(* IEC 61131-3 sources: plc-st-coding-agent/progress/evidence/f14_v14_remaining_20261113/jobs/custom_minimax-m27 (part 4) *)

(* ---- public-medium-02.raw_candidate_03.st ---- *)
TYPE ST_AnalogChannel :
STRUCT
    enable         : BOOL;
    hiLIM          : REAL;
    loLIM          : REAL;
    bipolar        : BOOL;
    measuringMode  : INT;
    retVal         : WORD;
    outputValue    : REAL;
END_STRUCT
END_TYPE;

FUNCTION_BLOCK FB_AnalogBatchProcessing
VAR_INPUT
    count : DINT;
END_VAR
VAR_IN_OUT
    analogValues : ARRAY[*] OF INT;
    channels     : ARRAY[*] OF ST_AnalogChannel;
END_VAR
VAR_OUTPUT
END_VAR
VAR
END_VAR

(*
ENGINEERING_CONTRACT
================================================================================
PUB001: Process 'count' channels starting at each array's lower bound.
        Arrays passed by reference preserve caller-defined bounds.
        Read-only: analogValues elements are never modified.
PUB002: Per-channel conversion based on measuringMode field.
        - Mode 0: Linear scaling using hiLIM/loLIM and bipolar flag.
        - Mode 1: Standard temperature (raw / 10.0).
        - Mode 2: Climatic temperature (raw / 100.0).
        - Invalid mode: retVal=16#8001, outputValue unchanged.
PUB003: Mode 0 linear scaling maps raw 0..27648 (unipolar) or -27648..27648 (bipolar)
        to loLIM..hiLIM range. OutputValue = loLIM + (raw - rawMin) * (hiLIM - loLIM) / range.
PUB004: If hiLIM <= loLIM in mode 0, set retVal=16#8002 and skip conversion.
PUB005: Disabled channels (enable=FALSE) are skipped; retVal and outputValue unchanged.
PUB006: Per-channel retVal WORD status: 16#8001 (invalid mode), 16#8002 (bad range).
PUB007: Same-scan priority: enable→measuringMode→hiLIM/loLIM check→conversion.
PUB008: Temperature output = raw / divisor (10 or 100) as REAL.
--------------------------------------------------------------------------------
*)

VAR
    tmpIndex     : DINT;
    tmpRaw       : INT;
    tmpRawReal   : REAL;
    tmpRange     : REAL;
    tmpOffset    : REAL;
    tmpChannel   : ST_AnalogChannel;
    tmpLower     : DINT;
    tmpUpperAna  : DINT;
    tmpUpperCh   : DINT;
    tmpProcessed : BOOL;
END_VAR

(* CONTRACT_RULES [] *)

tmpLower    := LOWER_BOUND(analogValues, 1);
tmpUpperAna := UPPER_BOUND(analogValues, 1);
tmpUpperCh  := UPPER_BOUND(channels, 1);

FOR tmpIndex := 0 TO (count - 1) DO
    tmpProcessed := FALSE;

    (* Bounds check: skip if index exceeds either array *)
    IF (tmpLower + tmpIndex) <= tmpUpperAna AND (tmpLower + tmpIndex) <= tmpUpperCh THEN
        tmpChannel := channels[tmpLower + tmpIndex];

        (* Skip disabled channels; retain previous outputValue and retVal *)
        IF tmpChannel.enable THEN

    (* Determine conversion based on measuringMode *)
    IF tmpChannel.measuringMode = 0 THEN
        (* Non-temperature linear scaling *)
        IF tmpChannel.hiLIM <= tmpChannel.loLIM THEN
            channels[tmpLower + tmpIndex].retVal := 16#8002;
        ELSE
            tmpRaw       := analogValues[tmpLower + tmpIndex];
            tmpRawReal   := TO_REAL(tmpRaw);
            tmpRange     := tmpChannel.hiLIM - tmpChannel.loLIM;

            IF tmpChannel.bipolar THEN
                (* Map -27648..27648 to loLIM..hiLIM *)
                tmpOffset    := TO_REAL(27648);
                channels[tmpLower + tmpIndex].outputValue := tmpChannel.loLIM +
                    (tmpRawReal + tmpOffset) * tmpRange / TO_REAL(55296);
            ELSE
                (* Map 0..27648 to loLIM..hiLIM *)
                channels[tmpLower + tmpIndex].outputValue := tmpChannel.loLIM +
                    tmpRawReal * tmpRange / TO_REAL(27648);
            END_IF;
            channels[tmpLower + tmpIndex].retVal := 0;
        END_IF;
        tmpProcessed := TRUE;
    ELSIF tmpChannel.measuringMode = 1 THEN
        (* Standard temperature: outputValue = raw / 10 *)
        tmpRaw := analogValues[tmpLower + tmpIndex];
        channels[tmpLower + tmpIndex].outputValue := TO_REAL(tmpRaw) / TO_REAL(10);
        channels[tmpLower + tmpIndex].retVal := 0;
        tmpProcessed := TRUE;
    ELSIF tmpChannel.measuringMode = 2 THEN
        (* Climatic temperature: outputValue = raw / 100 *)
        tmpRaw := analogValues[tmpLower + tmpIndex];
        channels[tmpLower + tmpIndex].outputValue := TO_REAL(tmpRaw) / TO_REAL(100);
        channels[tmpLower + tmpIndex].retVal := 0;
        tmpProcessed := TRUE;
    END_IF;

    (* Invalid measuringMode (not 0, 1, or 2) *)
    IF NOT tmpProcessed THEN
        channels[tmpLower + tmpIndex].retVal := 16#8001;
    END_IF;

    END_IF; (* close outer enable check *)

END_FOR;

END_FUNCTION_BLOCK

(* ---- public-medium-03.candidate_01.st ---- *)
FUNCTION_BLOCK FB_MovingAverage
VAR_INPUT
    cyclicExecution : BOOL;
    trigger         : BOOL;
    value           : LREAL;
    windowSize      : INT;
    reset           : BOOL;
END_VAR
VAR_OUTPUT
    average           : LREAL;
    windowSizeReached : BOOL;
    error             : BOOL;
    status            : WORD;
END_VAR
VAR
    circularBuffer : ARRAY[1..100] OF LREAL;
    bufferIndex    : INT := 1;
    sum             : LREAL := 0.0;
    sampleCount     : INT := 0;
    tmp_triggerPrev : BOOL := FALSE;
END_VAR
VAR_CONSTANT
    STATUS_OK           : WORD := 16#0000;
    STATUS_WINDOW_ERROR : WORD := 16#8200;
END_VAR

(*
ENGINEERING_CONTRACT
===================
Outputs and State Retention:
| Output/State        | Activation                    | Retention                  | Reset/Deactivation       | Same-scan Priority | Units/Boundaries     |
|---------------------|-------------------------------|----------------------------|--------------------------|--------------------| ---------------------|
| average             | New value added (cyclic/trig) | Held until next update     | reset=TRUE clears to 0.0 | cyclic>trigger     | LREAL, windowSize 1-100 |
| windowSizeReached   | sampleCount >= windowSize     | Held TRUE until reset      | reset=TRUE clears FALSE  | N/A                | BOOLEAN             |
| error               | windowSize<1 OR >100          | Held TRUE until valid/reset| reset=TRUE clears FALSE  | N/A                | BOOLEAN             |
| status              | Derived from error state      | Held until state change    | reset=TRUE clears to OK  | N/A                | WORD(16#0000/16#8200) |

Behavior:
- cyclicExecution=TRUE: add value every scan cycle (PUB001)
- trigger rising edge: add one value per press (PUB002)
- cyclicExecution has priority; trigger ignored when cyclic active
- reset clears buffer, sum, count, windowSizeReached (PUB003)
- Invalid windowSize (PUB004) sets error+status and halts processing
- windowSizeReached (PUB005): FALSE until window full, TRUE thereafter
- status codes (PUB006/PUB007): 16#0000=success, 16#8200=window error

First Scan: All VAR initializes to zero/false; no spurious trigger
Boundary: windowSize bounds [1,100] inclusive; strict comparison
)

(* CONTRACT_RULES [] *)

    // Rising edge detection for trigger
    IF trigger AND NOT tmp_triggerPrev THEN
        tmp_triggerPrev := trigger;
        IF NOT reset AND windowSize >= 1 AND windowSize <= 100 THEN
            // Buffer not yet full: add new value
            IF sampleCount < windowSize THEN
                sampleCount := sampleCount + 1;
                circularBuffer[sampleCount] := value;
                sum := sum + value;
                average := sum / TO_LREAL(sampleCount);
                IF sampleCount >= windowSize THEN
                    windowSizeReached := TRUE;
                END_IF;
            ELSE
                // Buffer full: replace oldest value using circular index
                sum := sum - circularBuffer[bufferIndex];
                circularBuffer[bufferIndex] := value;
                sum := sum + value;
                bufferIndex := (bufferIndex MOD windowSize) + 1;
                average := sum / TO_LREAL(windowSize);
            END_IF;
        END_IF;
    ELSE
        tmp_triggerPrev := trigger;
        // Check cyclicExecution on every scan when trigger not rising edge
        IF cyclicExecution AND NOT reset AND windowSize >= 1 AND windowSize <= 100 THEN
            // Buffer not yet full: add new value
            IF sampleCount < windowSize THEN
                sampleCount := sampleCount + 1;
                circularBuffer[sampleCount] := value;
                sum := sum + value;
                average := sum / TO_LREAL(sampleCount);
                IF sampleCount >= windowSize THEN
                    windowSizeReached := TRUE;
                END_IF;
            ELSE
                // Buffer full: replace oldest value using circular index
                sum := sum - circularBuffer[bufferIndex];
                circularBuffer[bufferIndex] := value;
                sum := sum + value;
                bufferIndex := (bufferIndex MOD windowSize) + 1;
                average := sum / TO_LREAL(windowSize);
            END_IF;
        END_IF;
    END_IF;

    // Reset handling - clears all state
    IF reset THEN
        bufferIndex := 1;
        sampleCount := 0;
        sum := 0.0;
        average := 0.0;
        windowSizeReached := FALSE;
        error := FALSE;
        status := STATUS_OK;
    ELSE
        // Validate window size when not resetting
        IF windowSize < 1 OR windowSize > 100 THEN
            error := TRUE;
            status := STATUS_WINDOW_ERROR;
        ELSE
            error := FALSE;
            status := STATUS_OK;
        END_IF;
    END_IF;

END_FUNCTION_BLOCK

(* ---- public-medium-03.candidate_02.st ---- *)
FUNCTION_BLOCK FB_MovingAverage
VAR_INPUT
    cyclicExecution : BOOL;
    trigger         : BOOL;
    value           : LREAL;
    windowSize      : INT;
    reset           : BOOL;
END_VAR
VAR_OUTPUT
    average           : LREAL;
    windowSizeReached : BOOL;
    error             : BOOL;
    status            : WORD;
END_VAR
VAR
    circularBuffer : ARRAY[1..100] OF LREAL;
    bufferIndex    : INT := 1;
    sum             : LREAL := 0.0;
    sampleCount     : INT := 0;
    tmp_triggerPrev : BOOL := FALSE;
END_VAR
VAR
    circularBuffer : ARRAY[1..100] OF LREAL;
    bufferIndex    : INT := 1;
    sum             : LREAL := 0.0;
    sampleCount     : INT := 0;
    tmp_triggerPrev : BOOL := FALSE;
END_VAR

(*
ENGINEERING_CONTRACT
===================
Outputs and State Retention:
| Output/State        | Activation                    | Retention                  | Reset/Deactivation       | Same-scan Priority | Units/Boundaries     |
|---------------------|-------------------------------|----------------------------|--------------------------|--------------------| ---------------------|
| average             | New value added (cyclic/trig) | Held until next update     | reset=TRUE clears to 0.0 | cyclic>trigger     | LREAL, windowSize 1-100 |
| windowSizeReached   | sampleCount >= windowSize     | Held TRUE until reset      | reset=TRUE clears FALSE  | N/A                | BOOLEAN             |
| error               | windowSize<1 OR >100          | Held TRUE until valid/reset| reset=TRUE clears FALSE  | N/A                | BOOLEAN             |
| status              | Derived from error state      | Held until state change    | reset=TRUE clears to OK  | N/A                | WORD(16#0000/16#8200) |

Behavior:
- cyclicExecution=TRUE: add value every scan cycle (PUB001)
- trigger rising edge: add one value per press (PUB002)
- cyclicExecution has priority; trigger ignored when cyclic active
- reset clears buffer, sum, count, windowSizeReached (PUB003)
- Invalid windowSize (PUB004) sets error+status and halts processing
- windowSizeReached (PUB005): FALSE until window full, TRUE thereafter
- status codes (PUB006/PUB007): 16#0000=success, 16#8200=window error

First Scan: All VAR initializes to zero/false; no spurious trigger
Boundary: windowSize bounds [1,100] inclusive; strict comparison
)

(* CONTRACT_RULES [] *)

    // Rising edge detection for trigger
    IF trigger AND NOT tmp_triggerPrev THEN
        tmp_triggerPrev := trigger;
        IF NOT reset AND windowSize >= 1 AND windowSize <= 100 THEN
            // Buffer not yet full: add new value
            IF sampleCount < windowSize THEN
                sampleCount := sampleCount + 1;
                circularBuffer[sampleCount] := value;
                sum := sum + value;
                average := sum / TO_LREAL(sampleCount);
                IF sampleCount >= windowSize THEN
                    windowSizeReached := TRUE;
                END_IF;
            ELSE
                // Buffer full: replace oldest value using circular index
                sum := sum - circularBuffer[bufferIndex];
                circularBuffer[bufferIndex] := value;
                sum := sum + value;
                bufferIndex := (bufferIndex MOD windowSize) + 1;
                average := sum / TO_LREAL(windowSize);
            END_IF;
        END_IF;
    ELSE
        tmp_triggerPrev := trigger;
        // Check cyclicExecution on every scan when trigger not rising edge
        IF cyclicExecution AND NOT reset AND windowSize >= 1 AND windowSize <= 100 THEN
            // Buffer not yet full: add new value
            IF sampleCount < windowSize THEN
                sampleCount := sampleCount + 1;
                circularBuffer[sampleCount] := value;
                sum := sum + value;
                average := sum / TO_LREAL(sampleCount);
                IF sampleCount >= windowSize THEN
                    windowSizeReached := TRUE;
                END_IF;
            ELSE
                // Buffer full: replace oldest value using circular index
                sum := sum - circularBuffer[bufferIndex];
                circularBuffer[bufferIndex] := value;
                sum := sum + value;
                bufferIndex := (bufferIndex MOD windowSize) + 1;
                average := sum / TO_LREAL(windowSize);
            END_IF;
        END_IF;
    END_IF;

    // Reset handling - clears all state
    IF reset THEN
        bufferIndex := 1;
        sampleCount := 0;
        sum := 0.0;
        average := 0.0;
        windowSizeReached := FALSE;
        error := FALSE;
        status := STATUS_OK;
    ELSE
        // Validate window size when not resetting
        IF windowSize < 1 OR windowSize > 100 THEN
            error := TRUE;
            status := STATUS_WINDOW_ERROR;
        ELSE
            error := FALSE;
            status := STATUS_OK;
        END_IF;
    END_IF;

END_FUNCTION_BLOCK

(* ---- public-medium-03.candidate_03.st ---- *)
FUNCTION_BLOCK FB_MovingAverage
VAR_INPUT
    cyclicExecution : BOOL;
    trigger         : BOOL;
    value           : LREAL;
    windowSize      : INT;
    reset           : BOOL;
END_VAR
VAR_OUTPUT
    average           : LREAL;
    windowSizeReached : BOOL;
    error             : BOOL;
    status            : WORD;
END_VAR
VAR
    circularBuffer : ARRAY[1..100] OF LREAL;
    bufferIndex    : INT := 1;
    sum             : LREAL := 0.0;
    sampleCount     : INT := 0;
    tmp_triggerPrev : BOOL := FALSE;
END_VAR

(*
ENGINEERING_CONTRACT
===================
Outputs and State Retention:
| Output/State        | Activation                    | Retention                  | Reset/Deactivation       | Same-scan Priority | Units/Boundaries     |
|---------------------|-------------------------------|----------------------------|--------------------------|--------------------| ---------------------|
| average             | New value added (cyclic/trig) | Held until next update     | reset=TRUE clears to 0.0 | cyclic>trigger     | LREAL, windowSize 1-100 |
| windowSizeReached   | sampleCount >= windowSize     | Held TRUE until reset      | reset=TRUE clears FALSE  | N/A                | BOOLEAN             |
| error               | windowSize<1 OR >100          | Held TRUE until valid/reset| reset=TRUE clears FALSE  | N/A                | BOOLEAN             |
| status              | Derived from error state      | Held until state change    | reset=TRUE clears to OK  | N/A                | WORD(16#0000/16#8200) |

Behavior:
- cyclicExecution=TRUE: add value every scan cycle (PUB001)
- trigger rising edge: add one value per press (PUB002)
- cyclicExecution has priority; trigger ignored when cyclic active
- reset clears buffer, sum, count, windowSizeReached (PUB003)
- Invalid windowSize (PUB004) sets error+status and halts processing
- windowSizeReached (PUB005): FALSE until window full, TRUE thereafter
- status codes (PUB006/PUB007): 16#0000=success, 16#8200=window error

First Scan: All VAR initializes to zero/false; no spurious trigger
Boundary: windowSize bounds [1,100] inclusive; strict comparison
*)

(* CONTRACT_RULES [] *)

    // Rising edge detection for trigger
    IF trigger AND NOT tmp_triggerPrev THEN
        tmp_triggerPrev := trigger;
        IF NOT reset AND windowSize >= 1 AND windowSize <= 100 THEN
            // Buffer not yet full: add new value
            IF sampleCount < windowSize THEN
                sampleCount := sampleCount + 1;
                circularBuffer[sampleCount] := value;
                sum := sum + value;
                average := sum / TO_LREAL(sampleCount);
                IF sampleCount >= windowSize THEN
                    windowSizeReached := TRUE;
                END_IF;
            ELSE
                // Buffer full: replace oldest value using circular index
                sum := sum - circularBuffer[bufferIndex];
                circularBuffer[bufferIndex] := value;
                sum := sum + value;
                bufferIndex := (bufferIndex MOD windowSize) + 1;
                average := sum / TO_LREAL(windowSize);
            END_IF;
        END_IF;
    ELSE
        tmp_triggerPrev := trigger;
        // Check cyclicExecution on every scan when trigger not rising edge
        IF cyclicExecution AND NOT reset AND windowSize >= 1 AND windowSize <= 100 THEN
            // Buffer not yet full: add new value
            IF sampleCount < windowSize THEN
                sampleCount := sampleCount + 1;
                circularBuffer[sampleCount] := value;
                sum := sum + value;
                average := sum / TO_LREAL(sampleCount);
                IF sampleCount >= windowSize THEN
                    windowSizeReached := TRUE;
                END_IF;
            ELSE
                // Buffer full: replace oldest value using circular index
                sum := sum - circularBuffer[bufferIndex];
                circularBuffer[bufferIndex] := value;
                sum := sum + value;
                bufferIndex := (bufferIndex MOD windowSize) + 1;
                average := sum / TO_LREAL(windowSize);
            END_IF;
        END_IF;
    END_IF;

    // Reset handling - clears all state
    IF reset THEN
        bufferIndex := 1;
        sampleCount := 0;
        sum := 0.0;
        average := 0.0;
        windowSizeReached := FALSE;
        error := FALSE;
        status := 16#0000;
    ELSE
        // Validate window size when not resetting
        IF windowSize < 1 OR windowSize > 100 THEN
            error := TRUE;
            status := 16#8200;
        ELSE
            error := FALSE;
            status := 16#0000;
        END_IF;
    END_IF;

END_FUNCTION_BLOCK

(* ---- public-medium-03.candidate_04.st ---- *)
FUNCTION_BLOCK FB_MovingAverage
VAR_INPUT
    cyclicExecution : BOOL;
    trigger         : BOOL;
    value           : LREAL;
    windowSize      : INT;
    reset           : BOOL;
END_VAR
VAR_OUTPUT
    average           : LREAL;
    windowSizeReached : BOOL;
    error             : BOOL;
    status            : WORD;
END_VAR
VAR
    circularBuffer    : ARRAY[1..100] OF LREAL;
    bufferIndex       : INT := 1;
    sum               : LREAL := 0.0;
    sampleCount       : INT := 0;
    tmp_triggerPrev   : BOOL := FALSE;
    tmp_windowSizePrev : INT := 0;
END_VAR

(*
ENGINEERING_CONTRACT
===================
Outputs and State Retention:
| Output/State        | Activation                    | Retention                  | Reset/Deactivation       | Same-scan Priority | Units/Boundaries     |
|---------------------|-------------------------------|----------------------------|--------------------------|--------------------| ---------------------|
| average             | New value added (cyclic/trig) | Held until next update     | reset=TRUE clears to 0.0 | cyclic>trigger     | LREAL, windowSize 1-100 |
| windowSizeReached   | sampleCount >= windowSize     | Held TRUE until reset      | reset=TRUE clears FALSE  | N/A                | BOOLEAN             |
| error               | windowSize<1 OR >100          | Held TRUE until valid/reset| reset=TRUE clears FALSE  | N/A                | BOOLEAN             |
| status              | Derived from error state      | Held until state change    | reset=TRUE clears to OK  | N/A                | WORD(16#0000/16#8200) |

Behavior:
- cyclicExecution=TRUE: add value every scan cycle (PUB001)
- trigger rising edge: add one value per press (PUB002)
- cyclicExecution has priority; trigger ignored when cyclic active
- reset clears buffer, sum, count, windowSizeReached (PUB003)
- Invalid windowSize (PUB004) sets error+status and halts processing
- windowSizeReached (PUB005): FALSE until window full, TRUE thereafter
- status codes (PUB006/PUB007): 16#0000=success, 16#8200=window error

First Scan: All VAR initializes to zero/false; no spurious trigger
Boundary: windowSize bounds [1,100] inclusive; strict comparison
*)

(* CONTRACT_RULES [] *)

    // Detect windowSize change and reset buffer state
    IF windowSize <> tmp_windowSizePrev THEN
        tmp_windowSizePrev := windowSize;
        FOR i := 1 TO 100 DO
            circularBuffer[i] := 0.0;
        END_FOR;
        bufferIndex := 1;
        sampleCount := 0;
        sum := 0.0;
    END_IF;

    // Rising edge detection for trigger takes priority over cyclicExecution
    IF trigger AND NOT tmp_triggerPrev THEN
        tmp_triggerPrev := trigger;
        IF NOT reset AND windowSize >= 1 AND windowSize <= 100 THEN
            // Buffer not yet full: add new value
            IF sampleCount < windowSize THEN
                sampleCount := sampleCount + 1;
                circularBuffer[sampleCount] := value;
                sum := sum + value;
                average := sum / TO_LREAL(sampleCount);
                IF sampleCount >= windowSize THEN
                    windowSizeReached := TRUE;
                END_IF;
            ELSE
                // Buffer full: replace oldest value using circular index
                sum := sum - circularBuffer[bufferIndex];
                circularBuffer[bufferIndex] := value;
                sum := sum + value;
                bufferIndex := (bufferIndex MOD windowSize) + 1;
                average := sum / TO_LREAL(windowSize);
            END_IF;
        END_IF;
    ELSIF cyclicExecution AND NOT tmp_triggerPrev THEN
        tmp_triggerPrev := trigger;
        // cyclicExecution every scan cycle when trigger not active
        IF NOT reset AND windowSize >= 1 AND windowSize <= 100 THEN
            // Buffer not yet full: add new value
            IF sampleCount < windowSize THEN
                sampleCount := sampleCount + 1;
                circularBuffer[sampleCount] := value;
                sum := sum + value;
                average := sum / TO_LREAL(sampleCount);
                IF sampleCount >= windowSize THEN
                    windowSizeReached := TRUE;
                END_IF;
            ELSE
                // Buffer full: replace oldest value using circular index
                sum := sum - circularBuffer[bufferIndex];
                circularBuffer[bufferIndex] := value;
                sum := sum + value;
                bufferIndex := (bufferIndex MOD windowSize) + 1;
                average := sum / TO_LREAL(windowSize);
            END_IF;
        END_IF;
    ELSE
        tmp_triggerPrev := trigger;
    END_IF;

    // Reset handling - clears all state
    IF reset THEN
        bufferIndex := 1;
        sampleCount := 0;
        sum := 0.0;
        average := 0.0;
        windowSizeReached := FALSE;
        error := FALSE;
        status := 16#0000;
    ELSE
        // Validate window size when not resetting
        IF windowSize < 1 OR windowSize > 100 THEN
            error := TRUE;
            status := 16#8200;
        ELSE
            error := FALSE;
            status := 16#0000;
        END_IF;
    END_IF;

END_FUNCTION_BLOCK

(* ---- public-medium-03.patch_base_02.st ---- *)
FUNCTION_BLOCK FB_MovingAverage
VAR_INPUT
    cyclicExecution : BOOL;
    trigger         : BOOL;
    value           : LREAL;
    windowSize      : INT;
    reset           : BOOL;
END_VAR
VAR_OUTPUT
    average           : LREAL;
    windowSizeReached : BOOL;
    error             : BOOL;
    status            : WORD;
END_VAR
VAR
    circularBuffer : ARRAY[1..100] OF LREAL;
    bufferIndex    : INT := 1;
    sum             : LREAL := 0.0;
    sampleCount     : INT := 0;
    tmp_triggerPrev : BOOL := FALSE;
END_VAR
VAR_CONSTANT
    STATUS_OK           : WORD := 16#0000;
    STATUS_WINDOW_ERROR : WORD := 16#8200;
END_VAR

(*
ENGINEERING_CONTRACT
===================
Outputs and State Retention:
| Output/State        | Activation                    | Retention                  | Reset/Deactivation       | Same-scan Priority | Units/Boundaries     |
|---------------------|-------------------------------|----------------------------|--------------------------|--------------------| ---------------------|
| average             | New value added (cyclic/trig) | Held until next update     | reset=TRUE clears to 0.0 | cyclic>trigger     | LREAL, windowSize 1-100 |
| windowSizeReached   | sampleCount >= windowSize     | Held TRUE until reset      | reset=TRUE clears FALSE  | N/A                | BOOLEAN             |
| error               | windowSize<1 OR >100          | Held TRUE until valid/reset| reset=TRUE clears FALSE  | N/A                | BOOLEAN             |
| status              | Derived from error state      | Held until state change    | reset=TRUE clears to OK  | N/A                | WORD(16#0000/16#8200) |

Behavior:
- cyclicExecution=TRUE: add value every scan cycle (PUB001)
- trigger rising edge: add one value per press (PUB002)
- cyclicExecution has priority; trigger ignored when cyclic active
- reset clears buffer, sum, count, windowSizeReached (PUB003)
- Invalid windowSize (PUB004) sets error+status and halts processing
- windowSizeReached (PUB005): FALSE until window full, TRUE thereafter
- status codes (PUB006/PUB007): 16#0000=success, 16#8200=window error

First Scan: All VAR initializes to zero/false; no spurious trigger
Boundary: windowSize bounds [1,100] inclusive; strict comparison
)

(* CONTRACT_RULES [] *)

    // Rising edge detection for trigger
    IF trigger AND NOT tmp_triggerPrev THEN
        tmp_triggerPrev := trigger;
        IF NOT reset AND windowSize >= 1 AND windowSize <= 100 THEN
            // Buffer not yet full: add new value
            IF sampleCount < windowSize THEN
                sampleCount := sampleCount + 1;
                circularBuffer[sampleCount] := value;
                sum := sum + value;
                average := sum / TO_LREAL(sampleCount);
                IF sampleCount >= windowSize THEN
                    windowSizeReached := TRUE;
                END_IF;
            ELSE
                // Buffer full: replace oldest value using circular index
                sum := sum - circularBuffer[bufferIndex];
                circularBuffer[bufferIndex] := value;
                sum := sum + value;
                bufferIndex := (bufferIndex MOD windowSize) + 1;
                average := sum / TO_LREAL(windowSize);
            END_IF;
        END_IF;
    ELSE
        tmp_triggerPrev := trigger;
        // Check cyclicExecution on every scan when trigger not rising edge
        IF cyclicExecution AND NOT reset AND windowSize >= 1 AND windowSize <= 100 THEN
            // Buffer not yet full: add new value
            IF sampleCount < windowSize THEN
                sampleCount := sampleCount + 1;
                circularBuffer[sampleCount] := value;
                sum := sum + value;
                average := sum / TO_LREAL(sampleCount);
                IF sampleCount >= windowSize THEN
                    windowSizeReached := TRUE;
                END_IF;
            ELSE
                // Buffer full: replace oldest value using circular index
                sum := sum - circularBuffer[bufferIndex];
                circularBuffer[bufferIndex] := value;
                sum := sum + value;
                bufferIndex := (bufferIndex MOD windowSize) + 1;
                average := sum / TO_LREAL(windowSize);
            END_IF;
        END_IF;
    END_IF;

    // Reset handling - clears all state
    IF reset THEN
        bufferIndex := 1;
        sampleCount := 0;
        sum := 0.0;
        average := 0.0;
        windowSizeReached := FALSE;
        error := FALSE;
        status := STATUS_OK;
    ELSE
        // Validate window size when not resetting
        IF windowSize < 1 OR windowSize > 100 THEN
            error := TRUE;
            status := STATUS_WINDOW_ERROR;
        ELSE
            error := FALSE;
            status := STATUS_OK;
        END_IF;
    END_IF;

END_FUNCTION_BLOCK

(* ---- public-medium-03.patch_base_03.st ---- *)
FUNCTION_BLOCK FB_MovingAverage
VAR_INPUT
    cyclicExecution : BOOL;
    trigger         : BOOL;
    value           : LREAL;
    windowSize      : INT;
    reset           : BOOL;
END_VAR
VAR_OUTPUT
    average           : LREAL;
    windowSizeReached : BOOL;
    error             : BOOL;
    status            : WORD;
END_VAR
VAR
    circularBuffer : ARRAY[1..100] OF LREAL;
    bufferIndex    : INT := 1;
    sum             : LREAL := 0.0;
    sampleCount     : INT := 0;
    tmp_triggerPrev : BOOL := FALSE;
END_VAR
VAR_CONSTANT
    STATUS_OK           : WORD := 16#0000;
    STATUS_WINDOW_ERROR : WORD := 16#8200;
END_VAR

(*
ENGINEERING_CONTRACT
===================
Outputs and State Retention:
| Output/State        | Activation                    | Retention                  | Reset/Deactivation       | Same-scan Priority | Units/Boundaries     |
|---------------------|-------------------------------|----------------------------|--------------------------|--------------------| ---------------------|
| average             | New value added (cyclic/trig) | Held until next update     | reset=TRUE clears to 0.0 | cyclic>trigger     | LREAL, windowSize 1-100 |
| windowSizeReached   | sampleCount >= windowSize     | Held TRUE until reset      | reset=TRUE clears FALSE  | N/A                | BOOLEAN             |
| error               | windowSize<1 OR >100          | Held TRUE until valid/reset| reset=TRUE clears FALSE  | N/A                | BOOLEAN             |
| status              | Derived from error state      | Held until state change    | reset=TRUE clears to OK  | N/A                | WORD(16#0000/16#8200) |

Behavior:
- cyclicExecution=TRUE: add value every scan cycle (PUB001)
- trigger rising edge: add one value per press (PUB002)
- cyclicExecution has priority; trigger ignored when cyclic active
- reset clears buffer, sum, count, windowSizeReached (PUB003)
- Invalid windowSize (PUB004) sets error+status and halts processing
- windowSizeReached (PUB005): FALSE until window full, TRUE thereafter
- status codes (PUB006/PUB007): 16#0000=success, 16#8200=window error

First Scan: All VAR initializes to zero/false; no spurious trigger
Boundary: windowSize bounds [1,100] inclusive; strict comparison
)

(* CONTRACT_RULES [] *)

    // Rising edge detection for trigger
    IF trigger AND NOT tmp_triggerPrev THEN
        tmp_triggerPrev := trigger;
        IF NOT reset AND windowSize >= 1 AND windowSize <= 100 THEN
            // Buffer not yet full: add new value
            IF sampleCount < windowSize THEN
                sampleCount := sampleCount + 1;
                circularBuffer[sampleCount] := value;
                sum := sum + value;
                average := sum / TO_LREAL(sampleCount);
                IF sampleCount >= windowSize THEN
                    windowSizeReached := TRUE;
                END_IF;
            ELSE
                // Buffer full: replace oldest value using circular index
                sum := sum - circularBuffer[bufferIndex];
                circularBuffer[bufferIndex] := value;
                sum := sum + value;
                bufferIndex := (bufferIndex MOD windowSize) + 1;
                average := sum / TO_LREAL(windowSize);
            END_IF;
        END_IF;
    ELSE
        tmp_triggerPrev := trigger;
        // Check cyclicExecution on every scan when trigger not rising edge
        IF cyclicExecution AND NOT reset AND windowSize >= 1 AND windowSize <= 100 THEN
            // Buffer not yet full: add new value
            IF sampleCount < windowSize THEN
                sampleCount := sampleCount + 1;
                circularBuffer[sampleCount] := value;
                sum := sum + value;
                average := sum / TO_LREAL(sampleCount);
                IF sampleCount >= windowSize THEN
                    windowSizeReached := TRUE;
                END_IF;
            ELSE
                // Buffer full: replace oldest value using circular index
                sum := sum - circularBuffer[bufferIndex];
                circularBuffer[bufferIndex] := value;
                sum := sum + value;
                bufferIndex := (bufferIndex MOD windowSize) + 1;
                average := sum / TO_LREAL(windowSize);
            END_IF;
        END_IF;
    END_IF;

    // Reset handling - clears all state
    IF reset THEN
        bufferIndex := 1;
        sampleCount := 0;
        sum := 0.0;
        average := 0.0;
        windowSizeReached := FALSE;
        error := FALSE;
        status := STATUS_OK;
    ELSE
        // Validate window size when not resetting
        IF windowSize < 1 OR windowSize > 100 THEN
            error := TRUE;
            status := STATUS_WINDOW_ERROR;
        ELSE
            error := FALSE;
            status := STATUS_OK;
        END_IF;
    END_IF;

END_FUNCTION_BLOCK

(* ---- public-medium-03.patch_base_04.st ---- *)
FUNCTION_BLOCK FB_MovingAverage
VAR_INPUT
    cyclicExecution : BOOL;
    trigger         : BOOL;
    value           : LREAL;
    windowSize      : INT;
    reset           : BOOL;
END_VAR
VAR_OUTPUT
    average           : LREAL;
    windowSizeReached : BOOL;
    error             : BOOL;
    status            : WORD;
END_VAR
VAR
    circularBuffer : ARRAY[1..100] OF LREAL;
    bufferIndex    : INT := 1;
    sum             : LREAL := 0.0;
    sampleCount     : INT := 0;
    tmp_triggerPrev : BOOL := FALSE;
END_VAR

(*
ENGINEERING_CONTRACT
===================
Outputs and State Retention:
| Output/State        | Activation                    | Retention                  | Reset/Deactivation       | Same-scan Priority | Units/Boundaries     |
|---------------------|-------------------------------|----------------------------|--------------------------|--------------------| ---------------------|
| average             | New value added (cyclic/trig) | Held until next update     | reset=TRUE clears to 0.0 | cyclic>trigger     | LREAL, windowSize 1-100 |
| windowSizeReached   | sampleCount >= windowSize     | Held TRUE until reset      | reset=TRUE clears FALSE  | N/A                | BOOLEAN             |
| error               | windowSize<1 OR >100          | Held TRUE until valid/reset| reset=TRUE clears FALSE  | N/A                | BOOLEAN             |
| status              | Derived from error state      | Held until state change    | reset=TRUE clears to OK  | N/A                | WORD(16#0000/16#8200) |

Behavior:
- cyclicExecution=TRUE: add value every scan cycle (PUB001)
- trigger rising edge: add one value per press (PUB002)
- cyclicExecution has priority; trigger ignored when cyclic active
- reset clears buffer, sum, count, windowSizeReached (PUB003)
- Invalid windowSize (PUB004) sets error+status and halts processing
- windowSizeReached (PUB005): FALSE until window full, TRUE thereafter
- status codes (PUB006/PUB007): 16#0000=success, 16#8200=window error

First Scan: All VAR initializes to zero/false; no spurious trigger
Boundary: windowSize bounds [1,100] inclusive; strict comparison
*)

(* CONTRACT_RULES [] *)

    // Rising edge detection for trigger
    IF trigger AND NOT tmp_triggerPrev THEN
        tmp_triggerPrev := trigger;
        IF NOT reset AND windowSize >= 1 AND windowSize <= 100 THEN
            // Buffer not yet full: add new value
            IF sampleCount < windowSize THEN
                sampleCount := sampleCount + 1;
                circularBuffer[sampleCount] := value;
                sum := sum + value;
                average := sum / TO_LREAL(sampleCount);
                IF sampleCount >= windowSize THEN
                    windowSizeReached := TRUE;
                END_IF;
            ELSE
                // Buffer full: replace oldest value using circular index
                sum := sum - circularBuffer[bufferIndex];
                circularBuffer[bufferIndex] := value;
                sum := sum + value;
                bufferIndex := (bufferIndex MOD windowSize) + 1;
                average := sum / TO_LREAL(windowSize);
            END_IF;
        END_IF;
    ELSE
        tmp_triggerPrev := trigger;
        // Check cyclicExecution on every scan when trigger not rising edge
        IF cyclicExecution AND NOT reset AND windowSize >= 1 AND windowSize <= 100 THEN
            // Buffer not yet full: add new value
            IF sampleCount < windowSize THEN
                sampleCount := sampleCount + 1;
                circularBuffer[sampleCount] := value;
                sum := sum + value;
                average := sum / TO_LREAL(sampleCount);
                IF sampleCount >= windowSize THEN
                    windowSizeReached := TRUE;
                END_IF;
            ELSE
                // Buffer full: replace oldest value using circular index
                sum := sum - circularBuffer[bufferIndex];
                circularBuffer[bufferIndex] := value;
                sum := sum + value;
                bufferIndex := (bufferIndex MOD windowSize) + 1;
                average := sum / TO_LREAL(windowSize);
            END_IF;
        END_IF;
    END_IF;

    // Reset handling - clears all state
    IF reset THEN
        bufferIndex := 1;
        sampleCount := 0;
        sum := 0.0;
        average := 0.0;
        windowSizeReached := FALSE;
        error := FALSE;
        status := 16#0000;
    ELSE
        // Validate window size when not resetting
        IF windowSize < 1 OR windowSize > 100 THEN
            error := TRUE;
            status := 16#8200;
        ELSE
            error := FALSE;
            status := 16#0000;
        END_IF;
    END_IF;

END_FUNCTION_BLOCK

(* ---- public-medium-03.raw_candidate_01.st ---- *)
FUNCTION_BLOCK FB_MovingAverage
VAR_INPUT
    cyclicExecution : BOOL;
    trigger         : BOOL;
    value           : LREAL;
    windowSize      : INT;
    reset           : BOOL;
END_VAR
VAR_OUTPUT
    average           : LREAL;
    windowSizeReached : BOOL;
    error             : BOOL;
    status            : WORD;
END_VAR
VAR
    circularBuffer : ARRAY[1..100] OF LREAL;
    bufferIndex    : INT := 1;
    sum             : LREAL := 0.0;
    sampleCount     : INT := 0;
    tmp_triggerPrev : BOOL := FALSE;
END_VAR
VAR_CONSTANT
    STATUS_OK           : WORD := 16#0000;
    STATUS_WINDOW_ERROR : WORD := 16#8200;
END_VAR

(*
ENGINEERING_CONTRACT
===================
Outputs and State Retention:
| Output/State        | Activation                    | Retention                  | Reset/Deactivation       | Same-scan Priority | Units/Boundaries     |
|---------------------|-------------------------------|----------------------------|--------------------------|--------------------| ---------------------|
| average             | New value added (cyclic/trig) | Held until next update     | reset=TRUE clears to 0.0 | cyclic>trigger     | LREAL, windowSize 1-100 |
| windowSizeReached   | sampleCount >= windowSize     | Held TRUE until reset      | reset=TRUE clears FALSE  | N/A                | BOOLEAN             |
| error               | windowSize<1 OR >100          | Held TRUE until valid/reset| reset=TRUE clears FALSE  | N/A                | BOOLEAN             |
| status              | Derived from error state      | Held until state change    | reset=TRUE clears to OK  | N/A                | WORD(16#0000/16#8200) |

Behavior:
- cyclicExecution=TRUE: add value every scan cycle (PUB001)
- trigger rising edge: add one value per press (PUB002)
- cyclicExecution has priority; trigger ignored when cyclic active
- reset clears buffer, sum, count, windowSizeReached (PUB003)
- Invalid windowSize (PUB004) sets error+status and halts processing
- windowSizeReached (PUB005): FALSE until window full, TRUE thereafter
- status codes (PUB006/PUB007): 16#0000=success, 16#8200=window error

First Scan: All VAR initializes to zero/false; no spurious trigger
Boundary: windowSize bounds [1,100] inclusive; strict comparison
)

(* CONTRACT_RULES [] *)

    // Rising edge detection for trigger
    IF trigger AND NOT tmp_triggerPrev THEN
        tmp_triggerPrev := trigger;
        IF NOT reset AND windowSize >= 1 AND windowSize <= 100 THEN
            // Buffer not yet full: add new value
            IF sampleCount < windowSize THEN
                sampleCount := sampleCount + 1;
                circularBuffer[sampleCount] := value;
                sum := sum + value;
                average := sum / TO_LREAL(sampleCount);
                IF sampleCount >= windowSize THEN
                    windowSizeReached := TRUE;
                END_IF;
            ELSE
                // Buffer full: replace oldest value using circular index
                sum := sum - circularBuffer[bufferIndex];
                circularBuffer[bufferIndex] := value;
                sum := sum + value;
                bufferIndex := (bufferIndex MOD windowSize) + 1;
                average := sum / TO_LREAL(windowSize);
            END_IF;
        END_IF;
    ELSE
        tmp_triggerPrev := trigger;
        // Check cyclicExecution on every scan when trigger not rising edge
        IF cyclicExecution AND NOT reset AND windowSize >= 1 AND windowSize <= 100 THEN
            // Buffer not yet full: add new value
            IF sampleCount < windowSize THEN
                sampleCount := sampleCount + 1;
                circularBuffer[sampleCount] := value;
                sum := sum + value;
                average := sum / TO_LREAL(sampleCount);
                IF sampleCount >= windowSize THEN
                    windowSizeReached := TRUE;
                END_IF;
            ELSE
                // Buffer full: replace oldest value using circular index
                sum := sum - circularBuffer[bufferIndex];
                circularBuffer[bufferIndex] := value;
                sum := sum + value;
                bufferIndex := (bufferIndex MOD windowSize) + 1;
                average := sum / TO_LREAL(windowSize);
            END_IF;
        END_IF;
    END_IF;

    // Reset handling - clears all state
    IF reset THEN
        bufferIndex := 1;
        sampleCount := 0;
        sum := 0.0;
        average := 0.0;
        windowSizeReached := FALSE;
        error := FALSE;
        status := STATUS_OK;
    ELSE
        // Validate window size when not resetting
        IF windowSize < 1 OR windowSize > 100 THEN
            error := TRUE;
            status := STATUS_WINDOW_ERROR;
        ELSE
            error := FALSE;
            status := STATUS_OK;
        END_IF;
    END_IF;

END_FUNCTION_BLOCK

(* ---- public-medium-03.raw_candidate_02.st ---- *)
FUNCTION_BLOCK FB_MovingAverage
VAR_INPUT
    cyclicExecution : BOOL;
    trigger         : BOOL;
    value           : LREAL;
    windowSize      : INT;
    reset           : BOOL;
END_VAR
VAR_OUTPUT
    average           : LREAL;
    windowSizeReached : BOOL;
    error             : BOOL;
    status            : WORD;
END_VAR
VAR
    circularBuffer : ARRAY[1..100] OF LREAL;
    bufferIndex    : INT := 1;
    sum             : LREAL := 0.0;
    sampleCount     : INT := 0;
    tmp_triggerPrev : BOOL := FALSE;
END_VAR
VAR
    circularBuffer : ARRAY[1..100] OF LREAL;
    bufferIndex    : INT := 1;
    sum             : LREAL := 0.0;
    sampleCount     : INT := 0;
    tmp_triggerPrev : BOOL := FALSE;
END_VAR

(*
ENGINEERING_CONTRACT
===================
Outputs and State Retention:
| Output/State        | Activation                    | Retention                  | Reset/Deactivation       | Same-scan Priority | Units/Boundaries     |
|---------------------|-------------------------------|----------------------------|--------------------------|--------------------| ---------------------|
| average             | New value added (cyclic/trig) | Held until next update     | reset=TRUE clears to 0.0 | cyclic>trigger     | LREAL, windowSize 1-100 |
| windowSizeReached   | sampleCount >= windowSize     | Held TRUE until reset      | reset=TRUE clears FALSE  | N/A                | BOOLEAN             |
| error               | windowSize<1 OR >100          | Held TRUE until valid/reset| reset=TRUE clears FALSE  | N/A                | BOOLEAN             |
| status              | Derived from error state      | Held until state change    | reset=TRUE clears to OK  | N/A                | WORD(16#0000/16#8200) |

Behavior:
- cyclicExecution=TRUE: add value every scan cycle (PUB001)
- trigger rising edge: add one value per press (PUB002)
- cyclicExecution has priority; trigger ignored when cyclic active
- reset clears buffer, sum, count, windowSizeReached (PUB003)
- Invalid windowSize (PUB004) sets error+status and halts processing
- windowSizeReached (PUB005): FALSE until window full, TRUE thereafter
- status codes (PUB006/PUB007): 16#0000=success, 16#8200=window error

First Scan: All VAR initializes to zero/false; no spurious trigger
Boundary: windowSize bounds [1,100] inclusive; strict comparison
)

(* CONTRACT_RULES [] *)

    // Rising edge detection for trigger
    IF trigger AND NOT tmp_triggerPrev THEN
        tmp_triggerPrev := trigger;
        IF NOT reset AND windowSize >= 1 AND windowSize <= 100 THEN
            // Buffer not yet full: add new value
            IF sampleCount < windowSize THEN
                sampleCount := sampleCount + 1;
                circularBuffer[sampleCount] := value;
                sum := sum + value;
                average := sum / TO_LREAL(sampleCount);
                IF sampleCount >= windowSize THEN
                    windowSizeReached := TRUE;
                END_IF;
            ELSE
                // Buffer full: replace oldest value using circular index
                sum := sum - circularBuffer[bufferIndex];
                circularBuffer[bufferIndex] := value;
                sum := sum + value;
                bufferIndex := (bufferIndex MOD windowSize) + 1;
                average := sum / TO_LREAL(windowSize);
            END_IF;
        END_IF;
    ELSE
        tmp_triggerPrev := trigger;
        // Check cyclicExecution on every scan when trigger not rising edge
        IF cyclicExecution AND NOT reset AND windowSize >= 1 AND windowSize <= 100 THEN
            // Buffer not yet full: add new value
            IF sampleCount < windowSize THEN
                sampleCount := sampleCount + 1;
                circularBuffer[sampleCount] := value;
                sum := sum + value;
                average := sum / TO_LREAL(sampleCount);
                IF sampleCount >= windowSize THEN
                    windowSizeReached := TRUE;
                END_IF;
            ELSE
                // Buffer full: replace oldest value using circular index
                sum := sum - circularBuffer[bufferIndex];
                circularBuffer[bufferIndex] := value;
                sum := sum + value;
                bufferIndex := (bufferIndex MOD windowSize) + 1;
                average := sum / TO_LREAL(windowSize);
            END_IF;
        END_IF;
    END_IF;

    // Reset handling - clears all state
    IF reset THEN
        bufferIndex := 1;
        sampleCount := 0;
        sum := 0.0;
        average := 0.0;
        windowSizeReached := FALSE;
        error := FALSE;
        status := STATUS_OK;
    ELSE
        // Validate window size when not resetting
        IF windowSize < 1 OR windowSize > 100 THEN
            error := TRUE;
            status := STATUS_WINDOW_ERROR;
        ELSE
            error := FALSE;
            status := STATUS_OK;
        END_IF;
    END_IF;

END_FUNCTION_BLOCK

(* ---- public-medium-03.raw_candidate_03.st ---- *)
FUNCTION_BLOCK FB_MovingAverage
VAR_INPUT
    cyclicExecution : BOOL;
    trigger         : BOOL;
    value           : LREAL;
    windowSize      : INT;
    reset           : BOOL;
END_VAR
VAR_OUTPUT
    average           : LREAL;
    windowSizeReached : BOOL;
    error             : BOOL;
    status            : WORD;
END_VAR
VAR
    circularBuffer : ARRAY[1..100] OF LREAL;
    bufferIndex    : INT := 1;
    sum             : LREAL := 0.0;
    sampleCount     : INT := 0;
    tmp_triggerPrev : BOOL := FALSE;
END_VAR

(*
ENGINEERING_CONTRACT
===================
Outputs and State Retention:
| Output/State        | Activation                    | Retention                  | Reset/Deactivation       | Same-scan Priority | Units/Boundaries     |
|---------------------|-------------------------------|----------------------------|--------------------------|--------------------| ---------------------|
| average             | New value added (cyclic/trig) | Held until next update     | reset=TRUE clears to 0.0 | cyclic>trigger     | LREAL, windowSize 1-100 |
| windowSizeReached   | sampleCount >= windowSize     | Held TRUE until reset      | reset=TRUE clears FALSE  | N/A                | BOOLEAN             |
| error               | windowSize<1 OR >100          | Held TRUE until valid/reset| reset=TRUE clears FALSE  | N/A                | BOOLEAN             |
| status              | Derived from error state      | Held until state change    | reset=TRUE clears to OK  | N/A                | WORD(16#0000/16#8200) |

Behavior:
- cyclicExecution=TRUE: add value every scan cycle (PUB001)
- trigger rising edge: add one value per press (PUB002)
- cyclicExecution has priority; trigger ignored when cyclic active
- reset clears buffer, sum, count, windowSizeReached (PUB003)
- Invalid windowSize (PUB004) sets error+status and halts processing
- windowSizeReached (PUB005): FALSE until window full, TRUE thereafter
- status codes (PUB006/PUB007): 16#0000=success, 16#8200=window error

First Scan: All VAR initializes to zero/false; no spurious trigger
Boundary: windowSize bounds [1,100] inclusive; strict comparison
*)

(* CONTRACT_RULES [] *)

    // Rising edge detection for trigger
    IF trigger AND NOT tmp_triggerPrev THEN
        tmp_triggerPrev := trigger;
        IF NOT reset AND windowSize >= 1 AND windowSize <= 100 THEN
            // Buffer not yet full: add new value
            IF sampleCount < windowSize THEN
                sampleCount := sampleCount + 1;
                circularBuffer[sampleCount] := value;
                sum := sum + value;
                average := sum / TO_LREAL(sampleCount);
                IF sampleCount >= windowSize THEN
                    windowSizeReached := TRUE;
                END_IF;
            ELSE
                // Buffer full: replace oldest value using circular index
                sum := sum - circularBuffer[bufferIndex];
                circularBuffer[bufferIndex] := value;
                sum := sum + value;
                bufferIndex := (bufferIndex MOD windowSize) + 1;
                average := sum / TO_LREAL(windowSize);
            END_IF;
        END_IF;
    ELSE
        tmp_triggerPrev := trigger;
        // Check cyclicExecution on every scan when trigger not rising edge
        IF cyclicExecution AND NOT reset AND windowSize >= 1 AND windowSize <= 100 THEN
            // Buffer not yet full: add new value
            IF sampleCount < windowSize THEN
                sampleCount := sampleCount + 1;
                circularBuffer[sampleCount] := value;
                sum := sum + value;
                average := sum / TO_LREAL(sampleCount);
                IF sampleCount >= windowSize THEN
                    windowSizeReached := TRUE;
                END_IF;
            ELSE
                // Buffer full: replace oldest value using circular index
                sum := sum - circularBuffer[bufferIndex];
                circularBuffer[bufferIndex] := value;
                sum := sum + value;
                bufferIndex := (bufferIndex MOD windowSize) + 1;
                average := sum / TO_LREAL(windowSize);
            END_IF;
        END_IF;
    END_IF;

    // Reset handling - clears all state
    IF reset THEN
        bufferIndex := 1;
        sampleCount := 0;
        sum := 0.0;
        average := 0.0;
        windowSizeReached := FALSE;
        error := FALSE;
        status := 16#0000;
    ELSE
        // Validate window size when not resetting
        IF windowSize < 1 OR windowSize > 100 THEN
            error := TRUE;
            status := 16#8200;
        ELSE
            error := FALSE;
            status := 16#0000;
        END_IF;
    END_IF;

END_FUNCTION_BLOCK

(* ---- public-medium-03.raw_candidate_04.st ---- *)
FUNCTION_BLOCK FB_MovingAverage
VAR_INPUT
    cyclicExecution : BOOL;
    trigger         : BOOL;
    value           : LREAL;
    windowSize      : INT;
    reset           : BOOL;
END_VAR
VAR_OUTPUT
    average           : LREAL;
    windowSizeReached : BOOL;
    error             : BOOL;
    status            : WORD;
END_VAR
VAR
    circularBuffer    : ARRAY[1..100] OF LREAL;
    bufferIndex       : INT := 1;
    sum               : LREAL := 0.0;
    sampleCount       : INT := 0;
    tmp_triggerPrev   : BOOL := FALSE;
    tmp_windowSizePrev : INT := 0;
END_VAR

(*
ENGINEERING_CONTRACT
===================
Outputs and State Retention:
| Output/State        | Activation                    | Retention                  | Reset/Deactivation       | Same-scan Priority | Units/Boundaries     |
|---------------------|-------------------------------|----------------------------|--------------------------|--------------------| ---------------------|
| average             | New value added (cyclic/trig) | Held until next update     | reset=TRUE clears to 0.0 | cyclic>trigger     | LREAL, windowSize 1-100 |
| windowSizeReached   | sampleCount >= windowSize     | Held TRUE until reset      | reset=TRUE clears FALSE  | N/A                | BOOLEAN             |
| error               | windowSize<1 OR >100          | Held TRUE until valid/reset| reset=TRUE clears FALSE  | N/A                | BOOLEAN             |
| status              | Derived from error state      | Held until state change    | reset=TRUE clears to OK  | N/A                | WORD(16#0000/16#8200) |

Behavior:
- cyclicExecution=TRUE: add value every scan cycle (PUB001)
- trigger rising edge: add one value per press (PUB002)
- cyclicExecution has priority; trigger ignored when cyclic active
- reset clears buffer, sum, count, windowSizeReached (PUB003)
- Invalid windowSize (PUB004) sets error+status and halts processing
- windowSizeReached (PUB005): FALSE until window full, TRUE thereafter
- status codes (PUB006/PUB007): 16#0000=success, 16#8200=window error

First Scan: All VAR initializes to zero/false; no spurious trigger
Boundary: windowSize bounds [1,100] inclusive; strict comparison
*)

(* CONTRACT_RULES [] *)

    // Detect windowSize change and reset buffer state
    IF windowSize <> tmp_windowSizePrev THEN
        tmp_windowSizePrev := windowSize;
        FOR i := 1 TO 100 DO
            circularBuffer[i] := 0.0;
        END_FOR;
        bufferIndex := 1;
        sampleCount := 0;
        sum := 0.0;
    END_IF;

    // Rising edge detection for trigger takes priority over cyclicExecution
    IF trigger AND NOT tmp_triggerPrev THEN
        tmp_triggerPrev := trigger;
        IF NOT reset AND windowSize >= 1 AND windowSize <= 100 THEN
            // Buffer not yet full: add new value
            IF sampleCount < windowSize THEN
                sampleCount := sampleCount + 1;
                circularBuffer[sampleCount] := value;
                sum := sum + value;
                average := sum / TO_LREAL(sampleCount);
                IF sampleCount >= windowSize THEN
                    windowSizeReached := TRUE;
                END_IF;
            ELSE
                // Buffer full: replace oldest value using circular index
                sum := sum - circularBuffer[bufferIndex];
                circularBuffer[bufferIndex] := value;
                sum := sum + value;
                bufferIndex := (bufferIndex MOD windowSize) + 1;
                average := sum / TO_LREAL(windowSize);
            END_IF;
        END_IF;
    ELSIF cyclicExecution AND NOT tmp_triggerPrev THEN
        tmp_triggerPrev := trigger;
        // cyclicExecution every scan cycle when trigger not active
        IF NOT reset AND windowSize >= 1 AND windowSize <= 100 THEN
            // Buffer not yet full: add new value
            IF sampleCount < windowSize THEN
                sampleCount := sampleCount + 1;
                circularBuffer[sampleCount] := value;
                sum := sum + value;
                average := sum / TO_LREAL(sampleCount);
                IF sampleCount >= windowSize THEN
                    windowSizeReached := TRUE;
                END_IF;
            ELSE
                // Buffer full: replace oldest value using circular index
                sum := sum - circularBuffer[bufferIndex];
                circularBuffer[bufferIndex] := value;
                sum := sum + value;
                bufferIndex := (bufferIndex MOD windowSize) + 1;
                average := sum / TO_LREAL(windowSize);
            END_IF;
        END_IF;
    ELSE
        tmp_triggerPrev := trigger;
    END_IF;

    // Reset handling - clears all state
    IF reset THEN
        bufferIndex := 1;
        sampleCount := 0;
        sum := 0.0;
        average := 0.0;
        windowSizeReached := FALSE;
        error := FALSE;
        status := 16#0000;
    ELSE
        // Validate window size when not resetting
        IF windowSize < 1 OR windowSize > 100 THEN
            error := TRUE;
            status := 16#8200;
        ELSE
            error := FALSE;
            status := 16#0000;
        END_IF;
    END_IF;

END_FUNCTION_BLOCK

(* ---- public-medium-04.candidate_01.st ---- *)
FUNCTION_BLOCK FB_TemperatureControl
VAR_INPUT
    TemperatureSensorInput : REAL;
    SetTemperature : REAL;
END_VAR
VAR_OUTPUT
    CurrentTemperature : REAL;
    SetTempDisplay : REAL;
    HeaterStatus : BOOL;
    OverheatProtection : BOOL;
    HeaterOutput : BOOL;
END_VAR
VAR
    OverheatTimer : TON;
    CooldownTimer : TON;
    tmp_SensorFault : BOOL;
END_VAR

(* ENGINEERING_CONTRACT:
 * | Output              | Activation                        | Retention/Hold              | Reset/Deactivation                    | Priority/Scan |
 * |---------------------|------------------------------------|-----------------------------|---------------------------------------|---------------|
 * | CurrentTemperature  | Every scan from sensor             | N/A (combinational read)    | N/A                                   | Same-scan     |
 * | SetTempDisplay      | Every scan from input              | N/A (combinational read)    | N/A                                   | Same-scan     |
 * | HeaterStatus        | Every scan = HeaterOutput          | N/A (combinational mirror)  | N/A                                   | Same-scan     |
 * | HeaterOutput        | Temp < SetTemp AND no fault/protection | Hold while conditions met | Sensor fault OR OverheatProtection OR Temp > SetTemp | Same-scan |
 * | OverheatProtection  | 5s continuous HeaterOutput         | Hold until 3s cooldown done | CooldownTimer.Q (elapsed >= 3s)       | Safety latch  |
 *
 * PUB001: HeaterOutput = (TemperatureSensorInput < SetTemperature) when no faults
 * PUB002, PUB005, PUB006, PUB008: Overheat triggers after TON.Q (elapsed >= 5s) with continuous heater ON
 *         3s cooldown via CooldownTimer before OverheatProtection can clear
 * PUB003: All status outputs updated every scan from current sensor/control state
 * PUB004: Sensor fault (temp < 0 OR temp > 100) disables heater immediately; no hysteresis on fault
 * Units: Temperature [degrees], Time [IEC TON with PT=T#5S/T#3S]
 *)

(* Initialize timers on first scan *)
OverheatTimer(IN := FALSE, PT := T#5S);
CooldownTimer(IN := FALSE, PT := T#3S);

(* PUB004: Sensor fault detection - immediate heater disable *)
tmp_SensorFault := (TemperatureSensorInput < 0.0) OR (TemperatureSensorInput > 100.0);

(* Primary control logic with safety priority *)
IF tmp_SensorFault THEN
    (* PUB004: Sensor fault - disable heater, enter protection state *)
    HeaterOutput := FALSE;
    OverheatProtection := TRUE;
    OverheatTimer(IN := FALSE);
    CooldownTimer(IN := TRUE, PT := T#3S);
    IF CooldownTimer.Q THEN
        OverheatProtection := FALSE;
        CooldownTimer(IN := FALSE);
    END_IF;

ELSIF OverheatProtection THEN
    (* PUB005, PUB008: Overheat protection active - heater forced OFF, cooldown in progress *)
    HeaterOutput := FALSE;
    CooldownTimer(IN := TRUE, PT := T#3S);
    OverheatTimer(IN := FALSE);
    IF CooldownTimer.Q THEN
        OverheatProtection := FALSE;
        CooldownTimer(IN := FALSE);
    END_IF;

ELSE
    (* Normal temperature control *)
    IF TemperatureSensorInput < SetTemperature THEN
        HeaterOutput := TRUE;
    ELSE
        HeaterOutput := FALSE;
    END_IF;

    (* PUB005, PUB006: Overheat protection - track 5s continuous heater operation *)
    IF HeaterOutput THEN
        OverheatTimer(IN := TRUE, PT := T#5S);
        IF OverheatTimer.Q THEN
            (* PUB002, PUB008: Overheat triggered - auto-off heater, start 3s cooldown *)
            OverheatProtection := TRUE;
            HeaterOutput := FALSE;
            OverheatTimer(IN := FALSE);
            CooldownTimer(IN := TRUE, PT := T#3S);
        END_IF;
    ELSE
        OverheatTimer(IN := FALSE);
    END_IF;
END_IF;

(* PUB003: Status display outputs updated every scan *)
CurrentTemperature := TemperatureSensorInput;
SetTempDisplay := SetTemperature;
HeaterStatus := HeaterOutput;
END_FUNCTION_BLOCK

(* CONTRACT_RULES [{"kind": "hold_until_reset", "output": "OverheatProtection", "set_input": null, "reset_input": null}] *)

(* ---- public-medium-04.patch_base_02.st ---- *)
FUNCTION_BLOCK FB_TemperatureControl
VAR_INPUT
    TemperatureSensorInput : REAL;
    SetTemperature : REAL;
END_VAR
VAR_OUTPUT
    CurrentTemperature : REAL;
    SetTempDisplay : REAL;
    HeaterStatus : BOOL;
    OverheatProtection : BOOL;
    HeaterOutput : BOOL;
END_VAR
VAR
    OverheatTimer : TON;
    CooldownTimer : TON;
    tmp_SensorFault : BOOL;
END_VAR

(* ENGINEERING_CONTRACT:
 * | Output              | Activation                        | Retention/Hold              | Reset/Deactivation                    | Priority/Scan |
 * |---------------------|------------------------------------|-----------------------------|---------------------------------------|---------------|
 * | CurrentTemperature  | Every scan from sensor             | N/A (combinational read)    | N/A                                   | Same-scan     |
 * | SetTempDisplay      | Every scan from input              | N/A (combinational read)    | N/A                                   | Same-scan     |
 * | HeaterStatus        | Every scan = HeaterOutput          | N/A (combinational mirror)  | N/A                                   | Same-scan     |
 * | HeaterOutput        | Temp < SetTemp AND no fault/protection | Hold while conditions met | Sensor fault OR OverheatProtection OR Temp > SetTemp | Same-scan |
 * | OverheatProtection  | 5s continuous HeaterOutput         | Hold until 3s cooldown done | CooldownTimer.Q (elapsed >= 3s)       | Safety latch  |
 *
 * PUB001: HeaterOutput = (TemperatureSensorInput < SetTemperature) when no faults
 * PUB002, PUB005, PUB006, PUB008: Overheat triggers after TON.Q (elapsed >= 5s) with continuous heater ON
 *         3s cooldown via CooldownTimer before OverheatProtection can clear
 * PUB003: All status outputs updated every scan from current sensor/control state
 * PUB004: Sensor fault (temp < 0 OR temp > 100) disables heater immediately; no hysteresis on fault
 * Units: Temperature [degrees], Time [IEC TON with PT=T#5S/T#3S]
 *)

(* Initialize timers on first scan *)
OverheatTimer(IN := FALSE, PT := T#5S);
CooldownTimer(IN := FALSE, PT := T#3S);

(* PUB004: Sensor fault detection - immediate heater disable *)
tmp_SensorFault := (TemperatureSensorInput < 0.0) OR (TemperatureSensorInput > 100.0);

(* Primary control logic with safety priority *)
IF tmp_SensorFault THEN
    (* PUB004: Sensor fault - disable heater, enter protection state *)
    HeaterOutput := FALSE;
    OverheatProtection := TRUE;
    OverheatTimer(IN := FALSE);
    CooldownTimer(IN := TRUE, PT := T#3S);
    IF CooldownTimer.Q THEN
        OverheatProtection := FALSE;
        CooldownTimer(IN := FALSE);
    END_IF;

ELSIF OverheatProtection THEN
    (* PUB005, PUB008: Overheat protection active - heater forced OFF, cooldown in progress *)
    HeaterOutput := FALSE;
    CooldownTimer(IN := TRUE, PT := T#3S);
    OverheatTimer(IN := FALSE);
    IF CooldownTimer.Q THEN
        OverheatProtection := FALSE;
        CooldownTimer(IN := FALSE);
    END_IF;

ELSE
    (* Normal temperature control *)
    IF TemperatureSensorInput < SetTemperature THEN
        HeaterOutput := TRUE;
    ELSE
        HeaterOutput := FALSE;
    END_IF;

    (* PUB005, PUB006: Overheat protection - track 5s continuous heater operation *)
    IF HeaterOutput THEN
        OverheatTimer(IN := TRUE, PT := T#5S);
        IF OverheatTimer.Q THEN
            (* PUB002, PUB008: Overheat triggered - auto-off heater, start 3s cooldown *)
            OverheatProtection := TRUE;
            HeaterOutput := FALSE;
            OverheatTimer(IN := FALSE);
            CooldownTimer(IN := TRUE, PT := T#3S);
        END_IF;
    ELSE
        OverheatTimer(IN := FALSE);
    END_IF;
END_IF;

(* PUB003: Status display outputs updated every scan *)
CurrentTemperature := TemperatureSensorInput;
SetTempDisplay := SetTemperature;
HeaterStatus := HeaterOutput;
END_FUNCTION_BLOCK

(* CONTRACT_RULES [{"kind": "hold_until_reset", "output": "OverheatProtection", "set_input": null, "reset_input": null}] *)

(* ---- public-medium-04.patch_base_03.st ---- *)
FUNCTION_BLOCK FB_TemperatureControl
VAR_INPUT
    TemperatureSensorInput : REAL;
    SetTemperature : REAL;
END_VAR
VAR_OUTPUT
    CurrentTemperature : REAL;
    SetTempDisplay : REAL;
    HeaterStatus : BOOL;
    OverheatProtection : BOOL;
    HeaterOutput : BOOL;
END_VAR
VAR
    OverheatTimer : TON;
    CooldownTimer : TON;
    tmp_SensorFault : BOOL;
END_VAR

(* ENGINEERING_CONTRACT:
 * | Output              | Activation                        | Retention/Hold              | Reset/Deactivation                    | Priority/Scan |
 * |---------------------|------------------------------------|-----------------------------|---------------------------------------|---------------|
 * | CurrentTemperature  | Every scan from sensor             | N/A (combinational read)    | N/A                                   | Same-scan     |
 * | SetTempDisplay      | Every scan from input              | N/A (combinational read)    | N/A                                   | Same-scan     |
 * | HeaterStatus        | Every scan = HeaterOutput          | N/A (combinational mirror)  | N/A                                   | Same-scan     |
 * | HeaterOutput        | Temp < SetTemp AND no fault/protection | Hold while conditions met | Sensor fault OR OverheatProtection OR Temp > SetTemp | Same-scan |
 * | OverheatProtection  | 5s continuous HeaterOutput         | Hold until 3s cooldown done | CooldownTimer.Q (elapsed >= 3s)       | Safety latch  |
 *
 * PUB001: HeaterOutput = (TemperatureSensorInput < SetTemperature) when no faults
 * PUB002, PUB005, PUB006, PUB008: Overheat triggers after TON.Q (elapsed >= 5s) with continuous heater ON
 *         3s cooldown via CooldownTimer before OverheatProtection can clear
 * PUB003: All status outputs updated every scan from current sensor/control state
 * PUB004: Sensor fault (temp < 0 OR temp > 100) disables heater immediately; no hysteresis on fault
 * Units: Temperature [degrees], Time [IEC TON with PT=T#5S/T#3S]
 *)

(* Initialize timers on first scan *)
OverheatTimer(IN := FALSE, PT := T#5S);
CooldownTimer(IN := FALSE, PT := T#3S);

(* PUB004: Sensor fault detection - immediate heater disable *)
tmp_SensorFault := (TemperatureSensorInput < 0.0) OR (TemperatureSensorInput > 100.0);

(* Primary control logic with safety priority *)
IF tmp_SensorFault THEN
    (* PUB004: Sensor fault - disable heater, enter protection state *)
    HeaterOutput := FALSE;
    OverheatProtection := TRUE;
    OverheatTimer(IN := FALSE);
    CooldownTimer(IN := TRUE, PT := T#3S);
    IF CooldownTimer.Q THEN
        OverheatProtection := FALSE;
        CooldownTimer(IN := FALSE);
    END_IF;

ELSIF OverheatProtection THEN
    (* PUB005, PUB008: Overheat protection active - heater forced OFF, cooldown in progress *)
    HeaterOutput := FALSE;
    CooldownTimer(IN := TRUE, PT := T#3S);
    OverheatTimer(IN := FALSE);
    IF CooldownTimer.Q THEN
        OverheatProtection := FALSE;
        CooldownTimer(IN := FALSE);
    END_IF;

ELSE
    (* Normal temperature control *)
    IF TemperatureSensorInput < SetTemperature THEN
        HeaterOutput := TRUE;
    ELSE
        HeaterOutput := FALSE;
    END_IF;

    (* PUB005, PUB006: Overheat protection - track 5s continuous heater operation *)
    IF HeaterOutput THEN
        OverheatTimer(IN := TRUE, PT := T#5S);
        IF OverheatTimer.Q THEN
            (* PUB002, PUB008: Overheat triggered - auto-off heater, start 3s cooldown *)
            OverheatProtection := TRUE;
            HeaterOutput := FALSE;
            OverheatTimer(IN := FALSE);
            CooldownTimer(IN := TRUE, PT := T#3S);
        END_IF;
    ELSE
        OverheatTimer(IN := FALSE);
    END_IF;
END_IF;

(* PUB003: Status display outputs updated every scan *)
CurrentTemperature := TemperatureSensorInput;
SetTempDisplay := SetTemperature;
HeaterStatus := HeaterOutput;
END_FUNCTION_BLOCK

(* CONTRACT_RULES [{"kind": "hold_until_reset", "output": "OverheatProtection", "set_input": null, "reset_input": null}] *)

(* ---- public-medium-04.raw_candidate_01.st ---- *)
FUNCTION_BLOCK FB_TemperatureControl
VAR_INPUT
    TemperatureSensorInput : REAL;
    SetTemperature : REAL;
END_VAR
VAR_OUTPUT
    CurrentTemperature : REAL;
    SetTempDisplay : REAL;
    HeaterStatus : BOOL;
    OverheatProtection : BOOL;
    HeaterOutput : BOOL;
END_VAR
VAR
    OverheatTimer : TON;
    CooldownTimer : TON;
    tmp_SensorFault : BOOL;
END_VAR

(* ENGINEERING_CONTRACT:
 * | Output              | Activation                        | Retention/Hold              | Reset/Deactivation                    | Priority/Scan |
 * |---------------------|------------------------------------|-----------------------------|---------------------------------------|---------------|
 * | CurrentTemperature  | Every scan from sensor             | N/A (combinational read)    | N/A                                   | Same-scan     |
 * | SetTempDisplay      | Every scan from input              | N/A (combinational read)    | N/A                                   | Same-scan     |
 * | HeaterStatus        | Every scan = HeaterOutput          | N/A (combinational mirror)  | N/A                                   | Same-scan     |
 * | HeaterOutput        | Temp < SetTemp AND no fault/protection | Hold while conditions met | Sensor fault OR OverheatProtection OR Temp > SetTemp | Same-scan |
 * | OverheatProtection  | 5s continuous HeaterOutput         | Hold until 3s cooldown done | CooldownTimer.Q (elapsed >= 3s)       | Safety latch  |
 *
 * PUB001: HeaterOutput = (TemperatureSensorInput < SetTemperature) when no faults
 * PUB002, PUB005, PUB006, PUB008: Overheat triggers after TON.Q (elapsed >= 5s) with continuous heater ON
 *         3s cooldown via CooldownTimer before OverheatProtection can clear
 * PUB003: All status outputs updated every scan from current sensor/control state
 * PUB004: Sensor fault (temp < 0 OR temp > 100) disables heater immediately; no hysteresis on fault
 * Units: Temperature [degrees], Time [IEC TON with PT=T#5S/T#3S]
 *)

(* Initialize timers on first scan *)
OverheatTimer(IN := FALSE, PT := T#5S);
CooldownTimer(IN := FALSE, PT := T#3S);

(* PUB004: Sensor fault detection - immediate heater disable *)
tmp_SensorFault := (TemperatureSensorInput < 0.0) OR (TemperatureSensorInput > 100.0);

(* Primary control logic with safety priority *)
IF tmp_SensorFault THEN
    (* PUB004: Sensor fault - disable heater, enter protection state *)
    HeaterOutput := FALSE;
    OverheatProtection := TRUE;
    OverheatTimer(IN := FALSE);
    CooldownTimer(IN := TRUE, PT := T#3S);
    IF CooldownTimer.Q THEN
        OverheatProtection := FALSE;
        CooldownTimer(IN := FALSE);
    END_IF;

ELSIF OverheatProtection THEN
    (* PUB005, PUB008: Overheat protection active - heater forced OFF, cooldown in progress *)
    HeaterOutput := FALSE;
    CooldownTimer(IN := TRUE, PT := T#3S);
    OverheatTimer(IN := FALSE);
    IF CooldownTimer.Q THEN
        OverheatProtection := FALSE;
        CooldownTimer(IN := FALSE);
    END_IF;

ELSE
    (* Normal temperature control *)
    IF TemperatureSensorInput < SetTemperature THEN
        HeaterOutput := TRUE;
    ELSE
        HeaterOutput := FALSE;
    END_IF;

    (* PUB005, PUB006: Overheat protection - track 5s continuous heater operation *)
    IF HeaterOutput THEN
        OverheatTimer(IN := TRUE, PT := T#5S);
        IF OverheatTimer.Q THEN
            (* PUB002, PUB008: Overheat triggered - auto-off heater, start 3s cooldown *)
            OverheatProtection := TRUE;
            HeaterOutput := FALSE;
            OverheatTimer(IN := FALSE);
            CooldownTimer(IN := TRUE, PT := T#3S);
        END_IF;
    ELSE
        OverheatTimer(IN := FALSE);
    END_IF;
END_IF;

(* PUB003: Status display outputs updated every scan *)
CurrentTemperature := TemperatureSensorInput;
SetTempDisplay := SetTemperature;
HeaterStatus := HeaterOutput;
END_FUNCTION_BLOCK

(* CONTRACT_RULES [{"kind": "hold_until_reset", "output": "OverheatProtection", "set_input": null, "reset_input": null}] *)

(* ---- public-medium-05.candidate_01.st ---- *)
(* ENGINEERING_CONTRACT
 * =============================================================================
 * Mode Switching (PUB001): Mode=0 manual, Mode=1 automatic. Output state on
 *   mode transition: both Motor outputs cleared, CompletionLight cleared.
 *   Transition detected via rising edge on Mode input variable.
 * Manual Mode (PUB002/PUB003):
 *   - Activation: Mode=0
 *   - Retention: MotorForward holds while ForwardButton=1 AND ReverseButton=0
 *   - Retention: MotorReverse holds while ReverseButton=1 AND ForwardButton=0
 *   - Deactivation: both cleared on any of: ForwardButton=0, ReverseButton=0,
 *     forward+reverse both asserted (interlock drops both), or Mode→1
 *   - Units: combinational, no timer
 * Automatic Mode (PUB004-PUB008):
 *   - Scan behavior: edge-sensitive state machine evaluated every scan
 *   - STATION_A activation: SensorA=TRUE AND State=IDLE
 *   - STATION_B activation: SensorB=TRUE AND State=MOVING_TO_B
 *   - STATION_C activation: SensorC=TRUE AND State=MOVING_TO_C
 *   - MotorForward activation: (State=IDLE AND SensorA=TRUE→ButtonA=TRUE)
 *     OR (State=STATION_A AND ButtonA=TRUE) OR (State=STATION_B AND ButtonB=TRUE)
 *   - MotorForward deactivation: on SensorB (→STATION_B) or SensorC (→STATION_C)
 *   - CompletionLight activation: SensorC=TRUE AND ButtonC=TRUE AND State=STATION_C
 *   - CompletionLight retention: holds until SensorC=FALSE (product removed)
 *   - CompletionLight deactivation: SensorC=FALSE transitions to IDLE
 *   - IDLE reset: State=IDLE when no product detected at any station
 *   - Units: boolean states, no timers
 * Same-scan priority: manual overrides automatic (Mode check first). Within
 *   automatic, state transition clears prior MotorForward before next sensor
 *   evaluation; CompletionLight set after Mode/state checks finalized.
 * Physical interlock: Pub002 prohibits MotorForward AND MotorReverse together.
 * =============================================================================
 *)

(* CONTRACT_RULES [] *)

FUNCTION_BLOCK ProductionLineControl
VAR_INPUT
    Mode            : BOOL;  (* 0=manual, 1=automatic *)
    ForwardButton   : BOOL;
    ReverseButton   : BOOL;
    SensorA         : BOOL;
    SensorB         : BOOL;
    SensorC         : BOOL;
    ButtonA         : BOOL;
    ButtonB         : BOOL;
    ButtonC         : BOOL;
END_VAR
VAR_OUTPUT
    MotorForward    : BOOL;
    MotorReverse    : BOOL;
    CompletionLight : BOOL;
END_VAR
VAR
    State           : INT;  (* 0=IDLE, 1=STATION_A, 2=MOVING_TO_B, 3=STATION_B,
                                4=MOVING_TO_C, 5=STATION_C *)
    tmp_PreviousMode : BOOL;
    tmp_ModeRising   : BOOL;
END_VAR

    (* Constants for state identification *)
    CONST
        IDLE         : INT := 0;
        STATION_A    : INT := 1;
        MOVING_TO_B  : INT := 2;
        STATION_B    : INT := 3;
        MOVING_TO_C  : INT := 4;
        STATION_C    : INT := 5;
    END_CONST

    (* Detect mode transition for reset behavior *)
    tmp_ModeRising := Mode AND NOT tmp_PreviousMode;
    tmp_PreviousMode := Mode;

    (* Reset outputs on mode entry into automatic *)
    IF tmp_ModeRising THEN
        MotorForward    := FALSE;
        MotorReverse    := FALSE;
        CompletionLight := FALSE;
    END_IF;

    (* Mode-based operation dispatch *)
    IF Mode = FALSE THEN
        (* Manual Mode (PUB002/PUB003) *)
        (* Interlock: forward and reverse cannot be energized together *)
        IF ForwardButton AND NOT ReverseButton THEN
            MotorForward := TRUE;
            MotorReverse := FALSE;
        ELSIF ReverseButton AND NOT ForwardButton THEN
            MotorForward := FALSE;
            MotorReverse := TRUE;
        ELSE
            MotorForward := FALSE;
            MotorReverse := FALSE;
        END_IF;
    ELSE
        (* Automatic Mode (PUB004-PUB008) *)
        MotorForward    := FALSE;
        MotorReverse    := FALSE;

        (* State machine evaluation *)
        CASE State OF
            IDLE :
                (* Wait for product at Workstation A *)
                IF SensorA THEN
                    State := STATION_A;
                END_IF;

            STATION_A :
                (* Product at Workstation A, wait for ButtonA *)
                IF ButtonA THEN
                    MotorForward := TRUE;
                    State := MOVING_TO_B;
                END_IF;
                (* Fallback: if product leaves A unexpectedly, return to IDLE *)
                IF NOT SensorA THEN
                    State := IDLE;
                END_IF;

            MOVING_TO_B :
                (* Motor running forward, wait for SensorB *)
                MotorForward := TRUE;
                IF SensorB THEN
                    MotorForward := FALSE;
                    State := STATION_B;
                END_IF;

            STATION_B :
                (* Product at Workstation B, wait for ButtonB *)
                IF ButtonB THEN
                    MotorForward := TRUE;
                    State := MOVING_TO_C;
                END_IF;
                (* Fallback: if product leaves B unexpectedly, return to IDLE *)
                IF NOT SensorB THEN
                    State := IDLE;
                END_IF;

            MOVING_TO_C :
                (* Motor running forward, wait for SensorC *)
                MotorForward := TRUE;
                IF SensorC THEN
                    MotorForward := FALSE;
                    State := STATION_C;
                END_IF;

            STATION_C :
                (* Product at Workstation C, wait for ButtonC, then product removal *)
                IF ButtonC THEN
                    CompletionLight := TRUE;
                END_IF;
                (* Product taken away: light off, return to IDLE *)
                IF NOT SensorC THEN
                    CompletionLight := FALSE;
                    State := IDLE;
                END_IF;

        END_CASE;
    END_IF;

END_FUNCTION_BLOCK

(* ---- public-medium-05.candidate_02.st ---- *)
TYPE ProductionState : INT (
    IDLE := 0,
    STATION_A := 1,
    MOVING_TO_B := 2,
    STATION_B := 3,
    MOVING_TO_C := 4,
    STATION_C := 5
);
END_TYPE;

(* ENGINEERING_CONTRACT
 * =============================================================================
 * Mode Switching (PUB001): Mode=0 manual, Mode=1 automatic. Output state on
 *   mode transition: both Motor outputs cleared, CompletionLight cleared.
 *   Transition detected via rising edge on Mode input variable.
 * Manual Mode (PUB002/PUB003):
 *   - Activation: Mode=0
 *   - Retention: MotorForward holds while ForwardButton=1 AND ReverseButton=0
 *   - Retention: MotorReverse holds while ReverseButton=1 AND ForwardButton=0
 *   - Deactivation: both cleared on any of: ForwardButton=0, ReverseButton=0,
 *     forward+reverse both asserted (interlock drops both), or Mode→1
 *   - Units: combinational, no timer
 * Automatic Mode (PUB004-PUB008):
 *   - Scan behavior: edge-sensitive state machine evaluated every scan
 *   - STATION_A activation: SensorA=TRUE AND State=IDLE
 *   - STATION_B activation: SensorB=TRUE AND State=MOVING_TO_B
 *   - STATION_C activation: SensorC=TRUE AND State=MOVING_TO_C
 *   - MotorForward activation: (State=IDLE AND SensorA=TRUE→ButtonA=TRUE)
 *     OR (State=STATION_A AND ButtonA=TRUE) OR (State=STATION_B AND ButtonB=TRUE)
 *   - MotorForward deactivation: on SensorB (→STATION_B) or SensorC (→STATION_C)
 *   - CompletionLight activation: SensorC=TRUE AND ButtonC=TRUE AND State=STATION_C
 *   - CompletionLight retention: holds until SensorC=FALSE (product removed)
 *   - CompletionLight deactivation: SensorC=FALSE transitions to IDLE
 *   - IDLE reset: State=IDLE when no product detected at any station
 *   - Units: boolean states, no timers
 * Same-scan priority: manual overrides automatic (Mode check first). Within
 *   automatic, state transition clears prior MotorForward before next sensor
 *   evaluation; CompletionLight set after Mode/state checks finalized.
 * Physical interlock: Pub002 prohibits MotorForward AND MotorReverse together.
 * =============================================================================
 *)

(* CONTRACT_RULES [] *)

FUNCTION_BLOCK ProductionLineControl
VAR_INPUT
    Mode            : BOOL;  (* 0=manual, 1=automatic *)
    ForwardButton   : BOOL;
    ReverseButton   : BOOL;
    SensorA         : BOOL;
    SensorB         : BOOL;
    SensorC         : BOOL;
    ButtonA         : BOOL;
    ButtonB         : BOOL;
    ButtonC         : BOOL;
END_VAR
VAR_OUTPUT
    MotorForward    : BOOL;
    MotorReverse    : BOOL;
    CompletionLight : BOOL;
END_VAR
VAR
    State           : INT;  (* 0=IDLE, 1=STATION_A, 2=MOVING_TO_B, 3=STATION_B,
                                4=MOVING_TO_C, 5=STATION_C *)
    tmp_PreviousMode : BOOL;
    tmp_ModeRising   : BOOL;
END_VAR

    (* Constants for state identification *)
    (* Detect mode transition for reset behavior *)
    tmp_ModeRising := Mode AND NOT tmp_PreviousMode;
    tmp_PreviousMode := Mode;

    (* Reset outputs on mode entry into automatic *)
    IF tmp_ModeRising THEN
        MotorForward    := FALSE;
        MotorReverse    := FALSE;
        CompletionLight := FALSE;
    END_IF;

    (* Mode-based operation dispatch *)
    IF Mode = FALSE THEN
        (* Manual Mode (PUB002/PUB003) *)
        (* Interlock: forward and reverse cannot be energized together *)
        IF ForwardButton AND NOT ReverseButton THEN
            MotorForward := TRUE;
            MotorReverse := FALSE;
        ELSIF ReverseButton AND NOT ForwardButton THEN
            MotorForward := FALSE;
            MotorReverse := TRUE;
        ELSE
            MotorForward := FALSE;
            MotorReverse := FALSE;
        END_IF;
    ELSE
        (* Automatic Mode (PUB004-PUB008) *)
        MotorForward    := FALSE;
        MotorReverse    := FALSE;

        (* State machine evaluation *)
        CASE State OF
            IDLE :
                (* Wait for product at Workstation A *)
                IF SensorA THEN
                    State := STATION_A;
                END_IF;

            STATION_A :
                (* Product at Workstation A, wait for ButtonA *)
                IF ButtonA THEN
                    MotorForward := TRUE;
                    State := MOVING_TO_B;
                END_IF;
                (* Fallback: if product leaves A unexpectedly, return to IDLE *)
                IF NOT SensorA THEN
                    State := IDLE;
                END_IF;

            MOVING_TO_B :
                (* Motor running forward, wait for SensorB *)
                MotorForward := TRUE;
                IF SensorB THEN
                    MotorForward := FALSE;
                    State := STATION_B;
                END_IF;

            STATION_B :
                (* Product at Workstation B, wait for ButtonB *)
                IF ButtonB THEN
                    MotorForward := TRUE;
                    State := MOVING_TO_C;
                END_IF;
                (* Fallback: if product leaves B unexpectedly, return to IDLE *)
                IF NOT SensorB THEN
                    State := IDLE;
                END_IF;

            MOVING_TO_C :
                (* Motor running forward, wait for SensorC *)
                MotorForward := TRUE;
                IF SensorC THEN
                    MotorForward := FALSE;
                    State := STATION_C;
                END_IF;

            STATION_C :
                (* Product at Workstation C, wait for ButtonC, then product removal *)
                IF ButtonC THEN
                    CompletionLight := TRUE;
                END_IF;
                (* Product taken away: light off, return to IDLE *)
                IF NOT SensorC THEN
                    CompletionLight := FALSE;
                    State := IDLE;
                END_IF;

        END_CASE;
    END_IF;

END_FUNCTION_BLOCK

(* ---- public-medium-05.candidate_03.st ---- *)
CONST
    IDLE         : INT := 0;
    STATION_A    : INT := 1;
    MOVING_TO_B  : INT := 2;
    STATION_B    : INT := 3;
    MOVING_TO_C  : INT := 4;
    STATION_C    : INT := 5;
END_CONST

(* ENGINEERING_CONTRACT
 * =============================================================================
 * Mode Switching (PUB001): Mode=0 manual, Mode=1 automatic. Output state on
 *   mode transition: both Motor outputs cleared, CompletionLight cleared.
 *   Transition detected via rising edge on Mode input variable.
 * Manual Mode (PUB002/PUB003):
 *   - Activation: Mode=0
 *   - Retention: MotorForward holds while ForwardButton=1 AND ReverseButton=0
 *   - Retention: MotorReverse holds while ReverseButton=1 AND ForwardButton=0
 *   - Deactivation: both cleared on any of: ForwardButton=0, ReverseButton=0,
 *     forward+reverse both asserted (interlock drops both), or Mode→1
 *   - Units: combinational, no timer
 * Automatic Mode (PUB004-PUB008):
 *   - Scan behavior: edge-sensitive state machine evaluated every scan
 *   - STATION_A activation: SensorA=TRUE AND State=IDLE
 *   - STATION_B activation: SensorB=TRUE AND State=MOVING_TO_B
 *   - STATION_C activation: SensorC=TRUE AND State=MOVING_TO_C
 *   - MotorForward activation: (State=IDLE AND SensorA=TRUE→ButtonA=TRUE)
 *     OR (State=STATION_A AND ButtonA=TRUE) OR (State=STATION_B AND ButtonB=TRUE)
 *   - MotorForward deactivation: on SensorB (→STATION_B) or SensorC (→STATION_C)
 *   - CompletionLight activation: SensorC=TRUE AND ButtonC=TRUE AND State=STATION_C
 *   - CompletionLight retention: holds until SensorC=FALSE (product removed)
 *   - CompletionLight deactivation: SensorC=FALSE transitions to IDLE
 *   - IDLE reset: State=IDLE when no product detected at any station
 *   - Units: boolean states, no timers
 * Same-scan priority: manual overrides automatic (Mode check first). Within
 *   automatic, state transition clears prior MotorForward before next sensor
 *   evaluation; CompletionLight set after Mode/state checks finalized.
 * Physical interlock: Pub002 prohibits MotorForward AND MotorReverse together.
 * =============================================================================
 *)

(* CONTRACT_RULES [] *)

FUNCTION_BLOCK ProductionLineControl
VAR_INPUT
    Mode            : BOOL;  (* 0=manual, 1=automatic *)
    ForwardButton   : BOOL;
    ReverseButton   : BOOL;
    SensorA         : BOOL;
    SensorB         : BOOL;
    SensorC         : BOOL;
    ButtonA         : BOOL;
    ButtonB         : BOOL;
    ButtonC         : BOOL;
END_VAR
VAR_OUTPUT
    MotorForward    : BOOL;
    MotorReverse    : BOOL;
    CompletionLight : BOOL;
END_VAR
VAR
    State           : INT;  (* 0=IDLE, 1=STATION_A, 2=MOVING_TO_B, 3=STATION_B,
                                4=MOVING_TO_C, 5=STATION_C *)
    tmp_PreviousMode : BOOL;
    tmp_ModeRising   : BOOL;
END_VAR

    (* Constants for state identification *)
    (* Detect mode transition for reset behavior *)
    tmp_ModeRising := Mode AND NOT tmp_PreviousMode;
    tmp_PreviousMode := Mode;

    (* Reset outputs on mode entry into automatic *)
    IF tmp_ModeRising THEN
        MotorForward    := FALSE;
        MotorReverse    := FALSE;
        CompletionLight := FALSE;
    END_IF;

    (* Mode-based operation dispatch *)
    IF Mode = FALSE THEN
        (* Manual Mode (PUB002/PUB003) *)
        (* Interlock: forward and reverse cannot be energized together *)
        IF ForwardButton AND NOT ReverseButton THEN
            MotorForward := TRUE;
            MotorReverse := FALSE;
        ELSIF ReverseButton AND NOT ForwardButton THEN
            MotorForward := FALSE;
            MotorReverse := TRUE;
        ELSE
            MotorForward := FALSE;
            MotorReverse := FALSE;
        END_IF;
    ELSE
        (* Automatic Mode (PUB004-PUB008) *)
        MotorForward    := FALSE;
        MotorReverse    := FALSE;

        (* State machine evaluation *)
        CASE State OF
            IDLE :
                (* Wait for product at Workstation A *)
                IF SensorA THEN
                    State := STATION_A;
                END_IF;

            STATION_A :
                (* Product at Workstation A, wait for ButtonA *)
                IF ButtonA THEN
                    MotorForward := TRUE;
                    State := MOVING_TO_B;
                END_IF;
                (* Fallback: if product leaves A unexpectedly, return to IDLE *)
                IF NOT SensorA THEN
                    State := IDLE;
                END_IF;

            MOVING_TO_B :
                (* Motor running forward, wait for SensorB *)
                MotorForward := TRUE;
                IF SensorB THEN
                    MotorForward := FALSE;
                    State := STATION_B;
                END_IF;

            STATION_B :
                (* Product at Workstation B, wait for ButtonB *)
                IF ButtonB THEN
                    MotorForward := TRUE;
                    State := MOVING_TO_C;
                END_IF;
                (* Fallback: if product leaves B unexpectedly, return to IDLE *)
                IF NOT SensorB THEN
                    State := IDLE;
                END_IF;

            MOVING_TO_C :
                (* Motor running forward, wait for SensorC *)
                MotorForward := TRUE;
                IF SensorC THEN
                    MotorForward := FALSE;
                    State := STATION_C;
                END_IF;

            STATION_C :
                (* Product at Workstation C, wait for ButtonC, then product removal *)
                IF ButtonC THEN
                    CompletionLight := TRUE;
                END_IF;
                (* Product taken away: light off, return to IDLE *)
                IF NOT SensorC THEN
                    CompletionLight := FALSE;
                    State := IDLE;
                END_IF;

        END_CASE;
    END_IF;

END_FUNCTION_BLOCK
